TYPE ST_PolarIIChamber_CtrlStatus EXTENDS ST_Module_CtrlStatus_Base :
STRUCT
	ServiceCtrl : ST_PolarIIChamber_ServiceCtrl;
	ServiceParam : ST_PolarIIChamber_ServiceParam;
	ServiceStatus : ST_PolarIIChamber_ServiceStatus;
END_STRUCT
END_TYPE

(* stored: Version 1.1.0.1, ProductVersion 3.1.4026.18
   DUT ST_PolarIIChamber_CtrlStatus: Id {14000000-0000-0000-0000-000000000076} *)
